(* IEC 61131-3 sources: Benedict-Informatik/Modul 319 Elektrotechnik/AND-Gatter_Test_mit_Visu, 1 file *)

(* ---- AND-Gatter_Test_mit_Visu_PLC_PRG.st ---- *)
PROGRAM PLC_PRG
VAR
	G3 : BOOL;
	G2 : BOOL;
	G1 : BOOL;
	M3 : BOOL;
	M1 : BOOL;
	M2 : BOOL;
END_VAR

(* Drei AND-Verknüpfungen mit je drei Eingängen *)
(* Achtung: Die Ausgänge sind teilweise ihre eigenen Eingänge und bleiben deshalb FALSE *)
G1 := M1 AND G2 AND G1;
G2 := M2 AND G1 AND G3;
G3 := M3 AND G3 AND G3;
